(* IEC 61131-3 sources: codesys-to-astra/tests/POUs/FB_C2aPid_Test, 5 files *)

(* ---- FB_C2aPid_Test.decl.st ---- *)
// Назначение: детерминированные свойства FB_C2aPid: ручной режим, ограничения выхода, знак П-звена.
//             Алгоритм ОВЕН STD_PID не повторяется (обёртка над Util.PID, исход check). Util.PID считает
//             по времени между вызовами, поэтому экземпляры живут в наборе, а проверка — через
//             CYCLES_TO_SETTLE циклов задачи.
// Автор:      kr0nsch
// Версия:     0.1.0
// Документ:   docs/TEST_REPORT.md
FUNCTION_BLOCK FB_C2aPid_Test EXTENDS coUnit.FB_TestSuite
VAR CONSTANT
    R_DELTA : REAL := 0.0001;       // допуск сравнения REAL
    CYCLES_TO_SETTLE : INT := 5;    // циклов до проверки
END_VAR
VAR
    fbManual : FB_C2aPid;   // ручной режим
    fbHigh : FB_C2aPid;     // насыщение сверху
    fbLow : FB_C2aPid;      // насыщение снизу
    fbSign : FB_C2aPid;     // знак П-звена
    iCycManual : INT;       // счётчик циклов теста ManualPassesThrough
    iCycHigh : INT;         // счётчик циклов теста OutputClampedHigh
    iCycLow : INT;          // счётчик циклов теста OutputClampedLow
    iCycSign : INT;         // счётчик циклов теста ProportionalSign
END_VAR

(* ---- ManualPassesThrough.method.impl.st ---- *)
coUnit.TEST('ManualPassesThrough');

fbManual(Y_MANUAL := 0.4, Y_MAN_SET := TRUE, PV := 10.0, SP := 50.0, XP := 10.0, TI := 0.0, TD := 0.0,
         PMIN := 0.0, PMAX := 1.0);
iCycManual := iCycManual + 1;
IF iCycManual >= CYCLES_TO_SETTLE THEN
    AssertEquals_REAL(Expected := 0.4, Actual := fbManual.Y, Delta := R_DELTA,
                      Message := CONCAT('manual, Y = ', REAL_TO_STRING(fbManual.Y)));
    coUnit.TEST_FINISHED();
END_IF

(* ---- OutputClampedHigh.method.impl.st ---- *)
coUnit.TEST('OutputClampedHigh');

fbHigh(PV := 0.0, SP := 1000.0, XP := 1.0, TI := 0.0, TD := 0.0, PMIN := 0.0, PMAX := 1.0);
iCycHigh := iCycHigh + 1;
IF iCycHigh >= CYCLES_TO_SETTLE THEN
    AssertEquals_REAL(Expected := 1.0, Actual := fbHigh.Y, Delta := R_DELTA,
                      Message := CONCAT('clamp high, Y = ', REAL_TO_STRING(fbHigh.Y)));
    coUnit.TEST_FINISHED();
END_IF

(* ---- OutputClampedLow.method.impl.st ---- *)
coUnit.TEST('OutputClampedLow');

fbLow(PV := 1000.0, SP := 0.0, XP := 1.0, TI := 0.0, TD := 0.0, PMIN := -0.5, PMAX := 1.0);
iCycLow := iCycLow + 1;
IF iCycLow >= CYCLES_TO_SETTLE THEN
    AssertEquals_REAL(Expected := -0.5, Actual := fbLow.Y, Delta := R_DELTA,
                      Message := CONCAT('clamp low, Y = ', REAL_TO_STRING(fbLow.Y)));
    coUnit.TEST_FINISHED();
END_IF

(* ---- ProportionalSign.method.impl.st ---- *)
coUnit.TEST('ProportionalSign');

fbSign(PV := 20.0, SP := 21.0, XP := 10.0, TI := 0.0, TD := 0.0, PMIN := -1.0, PMAX := 1.0);
iCycSign := iCycSign + 1;
IF iCycSign >= CYCLES_TO_SETTLE THEN
    AssertTrue(Condition := fbSign.Y > 0.0 AND fbSign.Y <= 1.0,
               Message := CONCAT('positive, Y = ', REAL_TO_STRING(fbSign.Y)));
    coUnit.TEST_FINISHED();
END_IF
